Universal Robots PolyScope program: Visor_easy_pick.urp

Program Visor_easy_pick (installation=default directory=/programs/02 Main Routines createdIn=5.19.0 lastSavedIn=5.19.0 robotSerialNumber=20245590068)
Calibrated DH parameters: a=[0.00013, -0.03651, -0.389144, 0.000102, 0.000008, 0]; d=[0.162613, 192.230671, -179.915756, -12.181517, 0.099698, 0.099535]; alpha=[1.57038, 0.002205, 0.004138, 1.570804, -1.571025, 0]; deltaTheta=[-0.000001, 1.484886, 4.928506, -0.130209, 0, 0]
InitVariablesNode variables(variable(name=easyPickCount_1, expression=0), variable(name=easyPickCount_2, expression=0), variable(name=easyPickNoObj_1, expression=0), variable(name=easyPickNoObj_2, expression=0), variable(name=easyPickParts_1, expression=0), variable(name=easyPickParts_2, expression=0))
Robot Program (runOnlyOnce=false)
  SafeHome (positionOptionType=SPEED_AND_ACCELERATION speed=1.047198 acceleration=1.396263 nextMotionTime=2)
  SuppressedNode
    MoveJ speed 60 deg/s, acceleration 80 deg/s^2 (useActiveTCP=true) feature=Base
      Waypoint Waypoint_1: TCP in base x=-394.49 y=66.162 z=300 mm, rx=0 ry=0 rz=-1.737 rad; joints [-170.007, -74.312, -107.466, -88.214, 90.137, -160.485] deg; TCP offset x=0 y=0 z=161 mm, rx=3.1415 ry=0 rz=0 rad
      Waypoint Waypoint_2: TCP in base x=-271.297 y=447.063 z=272.642 mm, rx=0.0644 ry=-0.0999 rz=-2.6762 rad; joints [-223.911, -95.236, -91.492, -88.214, 90.137, -160.485] deg
  SuppressedNode
    URCap VISOR Robotic App (SensoPart VISOR Robotic, SensoPart Industriesensorik GmbH) dataModel(visorAppTemplate=1); state(isChildrenLocked=true)
      URCap Easy Pick Setup (SensoPart VISOR Robotic, SensoPart Industriesensorik GmbH) dataModel(visorId=0, visorSetJob=true, visorJobName=Invite_table, visorImageAcqSetup=2, visorImageAcqSource=1, visorCalibSetNo=4, visorDetector=1, visorSetupStatus=5, visorOffsetSet=true, Pose(key=visorImageAcqPose, Position(key=posePosition, Length(key=X value=-0.259155 unit=M), Length(key=Y value=-0.466253 unit=M), Length(key=Z value=0.440005 unit=M)), Rotation(key=poseRotation, Angle(key=RX value=-0.000022 unit=RAD), Angle(key=RY value=-0.000009 unit=RAD), Angle(key=RZ value=-0.080607 unit=RAD))), Pose(key=visorGripPose, Position(key=posePosition, Length(key=X value=-0.331862 unit=M), Length(key=Y value=0.636112 unit=M), Length(key=Z value=-0.099161 unit=M)), Rotation(key=poseRotation, Angle(key=RX value=-0.000036 unit=RAD), Angle(key=RY value=0.000016 unit=RAD), Angle(key=RZ value=-3.091569 unit=RAD)))); state(isChildrenLocked=true)
      URCap Process (SensoPart VISOR Robotic, SensoPart Industriesensorik GmbH) dataModel(Variable(key=visorCounterVar, variable(name=easyPickCount, initializeExpression=0)), Variable(key=visorPartsFoundVar, variable(name=easyPickParts, initializeExpression=0))); state(isChildrenLocked=true)
        URCap Image Acquisition Pose (SensoPart VISOR Robotic, SensoPart Industriesensorik GmbH) state(isChildrenLocked=true)
        URCap Object Detected (SensoPart VISOR Robotic, SensoPart Industriesensorik GmbH) state(isChildrenLocked=true)
          Folder Open Gripper
            URCap Gripper (Robotiq_Grippers, Robotiq Inc.) dataModel(position=0.0, force=40.0, speed=26.0, positionInDouble=0.0, forceInDouble=40.0, speedInDouble=26.0, slaveIds=[9], blocking=true)
          URCap Approach Pose (SensoPart VISOR Robotic, SensoPart Industriesensorik GmbH) state(isChildrenLocked=true)
          URCap Target Pose (SensoPart VISOR Robotic, SensoPart Industriesensorik GmbH) state(isChildrenLocked=true)
          Folder Close Gripper
            URCap Gripper (Robotiq_Grippers, Robotiq Inc.) dataModel(position=30.19607843137255, force=40.0, speed=26.0, positionInDouble=30.19607843137255, forceInDouble=40.0, speedInDouble=26.0, slaveIds=[9], blocking=true)
          URCap Exit Pose (SensoPart VISOR Robotic, SensoPart Industriesensorik GmbH) state(isChildrenLocked=true)
        URCap No Object Detected (SensoPart VISOR Robotic, SensoPart Industriesensorik GmbH) dataModel(Variable(key=visorNoObjCountVar, variable(name=easyPickNoObj, initializeExpression=0)))
          Popup Message (haltProgram=false message=No object detected inputType=Text)
  SuppressedNode
    URCap VISOR Robotic App (SensoPart VISOR Robotic, SensoPart Industriesensorik GmbH) dataModel(visorAppTemplate=1); state(isChildrenLocked=true)
      URCap Easy Pick Setup (SensoPart VISOR Robotic, SensoPart Industriesensorik GmbH) dataModel(visorId=0, visorSetJob=true, visorImageAcqSetup=2, visorCalibSetNo=5, visorImageAcqSource=0, visorDetector=1, visorOffsetSet=true, visorJobName=Spatula_1, visorSetupStatus=3, Pose(key=visorGripPose, Position(key=posePosition, Length(key=X value=-0.690998 unit=M), Length(key=Y value=-0.162824 unit=M), Length(key=Z value=0.137826 unit=M)), Rotation(key=poseRotation, Angle(key=RX value=0.000034 unit=RAD), Angle(key=RY value=0.000118 unit=RAD), Angle(key=RZ value=-1.591974 unit=RAD))), Pose(key=visorImageAcqPose, Position(key=posePosition, Length(key=X value=-0.171937 unit=M), Length(key=Y value=-0.271355 unit=M), Length(key=Z value=0.185619 unit=M)), Rotation(key=poseRotation, Angle(key=RX value=-0.940927 unit=RAD), Angle(key=RY value=1.071665 unit=RAD), Angle(key=RZ value=-1.405061 unit=RAD)))); state(isChildrenLocked=true)
      URCap Process (SensoPart VISOR Robotic, SensoPart Industriesensorik GmbH) dataModel(Variable(key=visorCounterVar, variable(name=easyPickCount_1, initializeExpression=0)), Variable(key=visorPartsFoundVar, variable(name=easyPickParts_1, initializeExpression=0))); state(isChildrenLocked=true)
        URCap Image Acquisition Pose (SensoPart VISOR Robotic, SensoPart Industriesensorik GmbH) state(isChildrenLocked=true)
        URCap Object Detected (SensoPart VISOR Robotic, SensoPart Industriesensorik GmbH) state(isChildrenLocked=true)
          Folder Open Gripper
            URCap Gripper (Robotiq_Grippers, Robotiq Inc.) dataModel(position=43.13725490196078, force=0.0, speed=0.0, positionInDouble=43.13725490196078, forceInDouble=0.0, speedInDouble=0.0, slaveIds=[9], blocking=true)
            MoveJ speed 60 deg/s, acceleration 80 deg/s^2 (useActiveTCP=true) feature=Base
              Waypoint Waypoint_3: motionParameters(blendRadius=0.05); TCP in base x=-270.12 y=-355.427 z=307.888 mm, rx=0 ry=0 rz=2.3815 rad; joints [-109.801, -81.065, -101.124, -87.793, 90.132, 23.739] deg
              SuppressedNode
                Waypoint Waypoint_4: TCP in base x=-688.823 y=-159.742 z=166.597 mm, rx=0 ry=0.0001 rz=-1.6037 rad; joints [-155.999, -120.465, -74.71, -74.816, 90.152, -154.152] deg
          URCap Approach Pose (SensoPart VISOR Robotic, SensoPart Industriesensorik GmbH) dataModel(visorMotionType=1, visorOffsetZ=-25.0); state(isChildrenLocked=true)
          URCap Target Pose (SensoPart VISOR Robotic, SensoPart Industriesensorik GmbH) dataModel(visorToolSpeed=100.0, visorToolAcc=200.0); state(isChildrenLocked=true)
          Folder Close Gripper
            URCap Gripper (Robotiq_Grippers, Robotiq Inc.) dataModel(position=100.0, force=32.0, speed=34.0, positionInDouble=100.0, forceInDouble=32.0, speedInDouble=34.0, slaveIds=[9], blocking=true)
          URCap Exit Pose (SensoPart VISOR Robotic, SensoPart Industriesensorik GmbH) dataModel(visorToolSpeed=100.0, visorToolAcc=200.0, visorOffsetZ=-250.0); state(isChildrenLocked=true)
        URCap No Object Detected (SensoPart VISOR Robotic, SensoPart Industriesensorik GmbH) dataModel(Variable(key=visorNoObjCountVar, variable(name=easyPickNoObj_1, initializeExpression=0)))
          Popup Message (haltProgram=false message=No object inputType=Text)
  URCap VISOR Robotic App (SensoPart VISOR Robotic, SensoPart Industriesensorik GmbH) dataModel(visorAppTemplate=1); state(isChildrenLocked=true)
    URCap Easy Pick Setup (SensoPart VISOR Robotic, SensoPart Industriesensorik GmbH) dataModel(visorId=0, visorSetJob=true, visorJobName=Spatula_1, visorImageAcqSetup=2, visorCalibSetNo=6, visorDetector=1, visorImageAcqSource=1, visorOffsetSet=true, visorSetupStatus=5, Pose(key=visorImageAcqPose, Position(key=posePosition, Length(key=X value=-0.614958 unit=M), Length(key=Y value=-0.009338 unit=M), Length(key=Z value=0.311565 unit=M)), Rotation(key=poseRotation, Angle(key=RX value=0.00009 unit=RAD), Angle(key=RY value=0.000131 unit=RAD), Angle(key=RZ value=-1.603705 unit=RAD))), Pose(key=visorGripPose, Position(key=posePosition, Length(key=X value=-0.699816 unit=M), Length(key=Y value=-0.008571 unit=M), Length(key=Z value=-0.00748 unit=M)), Rotation(key=poseRotation, Angle(key=RX value=0.00001 unit=RAD), Angle(key=RY value=0.000002 unit=RAD), Angle(key=RZ value=-1.551141 unit=RAD)))); state(isChildrenLocked=true)
    URCap Process (SensoPart VISOR Robotic, SensoPart Industriesensorik GmbH) dataModel(Variable(key=visorCounterVar, variable(name=easyPickCount_2, initializeExpression=0)), Variable(key=visorPartsFoundVar, variable(name=easyPickParts_2, initializeExpression=0))); state(isChildrenLocked=true)
      URCap Image Acquisition Pose (SensoPart VISOR Robotic, SensoPart Industriesensorik GmbH) state(isChildrenLocked=true)
      URCap Object Detected (SensoPart VISOR Robotic, SensoPart Industriesensorik GmbH) state(isChildrenLocked=true)
        Folder Open Gripper
          URCap Gripper (Robotiq_Grippers, Robotiq Inc.) dataModel(position=24.705882352941178, force=30.19607843137255, speed=36.07843137254902, positionInDouble=24.705882352941178, forceInDouble=30.19607843137255, speedInDouble=36.07843137254902, slaveIds=[9], blocking=true)
        URCap Approach Pose (SensoPart VISOR Robotic, SensoPart Industriesensorik GmbH) dataModel(visorOffsetZ=-70.0); state(isChildrenLocked=true)
        URCap Target Pose (SensoPart VISOR Robotic, SensoPart Industriesensorik GmbH) dataModel(visorOffsetZ=0.0); state(isChildrenLocked=true)
        Folder Close Gripper
          URCap Gripper (Robotiq_Grippers, Robotiq Inc.) dataModel(position=100.0, force=30.19607843137255, speed=36.07843137254902, positionInDouble=100.0, forceInDouble=30.19607843137255, speedInDouble=36.07843137254902, slaveIds=[9], blocking=true)
        URCap Exit Pose (SensoPart VISOR Robotic, SensoPart Industriesensorik GmbH) dataModel(visorOffsetZ=0.0); state(isChildrenLocked=true)
      URCap No Object Detected (SensoPart VISOR Robotic, SensoPart Industriesensorik GmbH) dataModel(Variable(key=visorNoObjCountVar, variable(name=easyPickNoObj_2, initializeExpression=0)))
        Popup Message (haltProgram=false message=No object detected inputType=Text)
  MoveJ speed 60 deg/s, acceleration 80 deg/s^2 (useActiveTCP=true) feature=Base
    Waypoint Waypoint_5: TCP in base x=-503.981 y=-20.518 z=-8.277 mm, rx=0 ry=0 rz=-1.552 rad; joints [-162.341, -110.08, -122.165, -37.748, 90.081, -163.302] deg
    Waypoint Waypoint_6: TCP in base x=-503.981 y=-20.518 z=254.365 mm, rx=0 ry=0 rz=-1.552 rad; joints [-162.295, -90.141, -100.676, -79.176, 90.138, -163.366] deg
  SafeHome (positionOptionType=SPEED_AND_ACCELERATION speed=1.047198 acceleration=1.396263 nextMotionTime=2)
  URCap Gripper (Robotiq_Grippers, Robotiq Inc.) dataModel(position=0.0, force=30.19607843137255, speed=36.07843137254902, positionInDouble=0.0, forceInDouble=30.19607843137255, speedInDouble=36.07843137254902, slaveIds=[9], blocking=true)
